FUNCTION_BLOCK SortingRouteConditions (* Sorting-only architecture following Distribution and tutorial modules 1-4 *)
  (* Standard: 61499-2 *)
  (* Version 2.0, 2026-11-09, sorting2n, sorting2n *)
  PACKAGE Main;
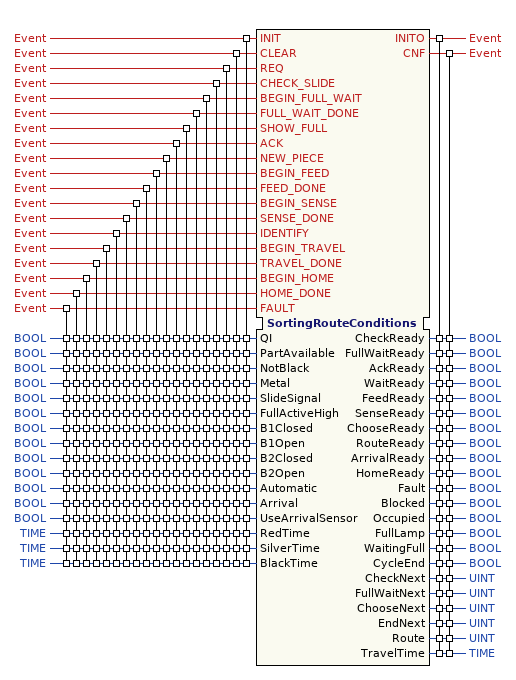
  EVENT_INPUT
    INIT WITH QI, PartAvailable, NotBlack, Metal, SlideSignal, FullActiveHigh, B1Closed, B1Open, B2Closed, B2Open, Automatic, Arrival, UseArrivalSensor, RedTime, SilverTime, BlackTime;
    CLEAR WITH QI, PartAvailable, NotBlack, Metal, SlideSignal, FullActiveHigh, B1Closed, B1Open, B2Closed, B2Open, Automatic, Arrival, UseArrivalSensor, RedTime, SilverTime, BlackTime;
    REQ WITH QI, PartAvailable, NotBlack, Metal, SlideSignal, FullActiveHigh, B1Closed, B1Open, B2Closed, B2Open, Automatic, Arrival, UseArrivalSensor, RedTime, SilverTime, BlackTime;
    CHECK_SLIDE WITH QI, PartAvailable, NotBlack, Metal, SlideSignal, FullActiveHigh, B1Closed, B1Open, B2Closed, B2Open, Automatic, Arrival, UseArrivalSensor, RedTime, SilverTime, BlackTime;
    BEGIN_FULL_WAIT WITH QI, PartAvailable, NotBlack, Metal, SlideSignal, FullActiveHigh, B1Closed, B1Open, B2Closed, B2Open, Automatic, Arrival, UseArrivalSensor, RedTime, SilverTime, BlackTime;
    FULL_WAIT_DONE WITH QI, PartAvailable, NotBlack, Metal, SlideSignal, FullActiveHigh, B1Closed, B1Open, B2Closed, B2Open, Automatic, Arrival, UseArrivalSensor, RedTime, SilverTime, BlackTime;
    SHOW_FULL WITH QI, PartAvailable, NotBlack, Metal, SlideSignal, FullActiveHigh, B1Closed, B1Open, B2Closed, B2Open, Automatic, Arrival, UseArrivalSensor, RedTime, SilverTime, BlackTime;
    ACK WITH QI, PartAvailable, NotBlack, Metal, SlideSignal, FullActiveHigh, B1Closed, B1Open, B2Closed, B2Open, Automatic, Arrival, UseArrivalSensor, RedTime, SilverTime, BlackTime;
    NEW_PIECE WITH QI, PartAvailable, NotBlack, Metal, SlideSignal, FullActiveHigh, B1Closed, B1Open, B2Closed, B2Open, Automatic, Arrival, UseArrivalSensor, RedTime, SilverTime, BlackTime;
    BEGIN_FEED WITH QI, PartAvailable, NotBlack, Metal, SlideSignal, FullActiveHigh, B1Closed, B1Open, B2Closed, B2Open, Automatic, Arrival, UseArrivalSensor, RedTime, SilverTime, BlackTime;
    FEED_DONE WITH QI, PartAvailable, NotBlack, Metal, SlideSignal, FullActiveHigh, B1Closed, B1Open, B2Closed, B2Open, Automatic, Arrival, UseArrivalSensor, RedTime, SilverTime, BlackTime;
    BEGIN_SENSE WITH QI, PartAvailable, NotBlack, Metal, SlideSignal, FullActiveHigh, B1Closed, B1Open, B2Closed, B2Open, Automatic, Arrival, UseArrivalSensor, RedTime, SilverTime, BlackTime;
    SENSE_DONE WITH QI, PartAvailable, NotBlack, Metal, SlideSignal, FullActiveHigh, B1Closed, B1Open, B2Closed, B2Open, Automatic, Arrival, UseArrivalSensor, RedTime, SilverTime, BlackTime;
    IDENTIFY WITH QI, PartAvailable, NotBlack, Metal, SlideSignal, FullActiveHigh, B1Closed, B1Open, B2Closed, B2Open, Automatic, Arrival, UseArrivalSensor, RedTime, SilverTime, BlackTime;
    BEGIN_TRAVEL WITH QI, PartAvailable, NotBlack, Metal, SlideSignal, FullActiveHigh, B1Closed, B1Open, B2Closed, B2Open, Automatic, Arrival, UseArrivalSensor, RedTime, SilverTime, BlackTime;
    TRAVEL_DONE WITH QI, PartAvailable, NotBlack, Metal, SlideSignal, FullActiveHigh, B1Closed, B1Open, B2Closed, B2Open, Automatic, Arrival, UseArrivalSensor, RedTime, SilverTime, BlackTime;
    BEGIN_HOME WITH QI, PartAvailable, NotBlack, Metal, SlideSignal, FullActiveHigh, B1Closed, B1Open, B2Closed, B2Open, Automatic, Arrival, UseArrivalSensor, RedTime, SilverTime, BlackTime;
    HOME_DONE WITH QI, PartAvailable, NotBlack, Metal, SlideSignal, FullActiveHigh, B1Closed, B1Open, B2Closed, B2Open, Automatic, Arrival, UseArrivalSensor, RedTime, SilverTime, BlackTime;
    FAULT WITH QI, PartAvailable, NotBlack, Metal, SlideSignal, FullActiveHigh, B1Closed, B1Open, B2Closed, B2Open, Automatic, Arrival, UseArrivalSensor, RedTime, SilverTime, BlackTime;
  END_EVENT
  EVENT_OUTPUT
    INITO WITH CheckReady, FullWaitReady, AckReady, WaitReady, FeedReady, SenseReady, ChooseReady, RouteReady, ArrivalReady, HomeReady, Fault, Blocked, Occupied, FullLamp, WaitingFull, CycleEnd, CheckNext, FullWaitNext, ChooseNext, EndNext, Route, TravelTime;
    CNF WITH CheckReady, FullWaitReady, AckReady, WaitReady, FeedReady, SenseReady, ChooseReady, RouteReady, ArrivalReady, HomeReady, Fault, Blocked, Occupied, FullLamp, WaitingFull, CycleEnd, CheckNext, FullWaitNext, ChooseNext, EndNext, Route, TravelTime;
  END_EVENT
  VAR_INPUT
    QI : BOOL := FALSE;
    PartAvailable : BOOL := FALSE;
    NotBlack : BOOL := FALSE;
    Metal : BOOL := FALSE;
    SlideSignal : BOOL := FALSE;
    FullActiveHigh : BOOL := FALSE;
    B1Closed : BOOL := FALSE;
    B1Open : BOOL := FALSE;
    B2Closed : BOOL := FALSE;
    B2Open : BOOL := FALSE;
    Automatic : BOOL := FALSE;
    Arrival : BOOL := FALSE;
    UseArrivalSensor : BOOL := FALSE;
    RedTime : TIME := T#2500ms;
    SilverTime : TIME := T#3s;
    BlackTime : TIME := T#5s;
  END_VAR
  VAR_OUTPUT
    CheckReady : BOOL := FALSE;
    FullWaitReady : BOOL := FALSE;
    AckReady : BOOL := FALSE;
    WaitReady : BOOL := FALSE;
    FeedReady : BOOL := FALSE;
    SenseReady : BOOL := FALSE;
    ChooseReady : BOOL := FALSE;
    RouteReady : BOOL := FALSE;
    ArrivalReady : BOOL := FALSE;
    HomeReady : BOOL := FALSE;
    Fault : BOOL := FALSE;
    Blocked : BOOL := FALSE;
    Occupied : BOOL := FALSE;
    FullLamp : BOOL := FALSE;
    WaitingFull : BOOL := FALSE;
    CycleEnd : BOOL := FALSE;
    CheckNext : UINT := 0;
    FullWaitNext : UINT := 0;
    ChooseNext : UINT := 0;
    EndNext : UINT := 0;
    Route : UINT := 0;
    TravelTime : TIME := T#5s;
  END_VAR
  VAR
    FeedElapsed : BOOL;
    SenseElapsed : BOOL;
    FinishElapsed : BOOL;
    TravelElapsed : BOOL;
    HomeElapsed : BOOL;
    Acked : BOOL;
  END_VAR
  EC_STATES
    IDLE;
    ON_INIT : ON_INIT -> INITO;
    ON_CLEAR : ON_CLEAR -> CNF;
    ON_REQ : ON_REQ -> CNF;
    ON_CHECK_SLIDE : ON_CHECK_SLIDE -> CNF;
    ON_BEGIN_FULL_WAIT : ON_BEGIN_FULL_WAIT -> CNF;
    ON_FULL_WAIT_DONE : ON_FULL_WAIT_DONE -> CNF;
    ON_SHOW_FULL : ON_SHOW_FULL -> CNF;
    ON_ACK : ON_ACK -> CNF;
    ON_NEW_PIECE : ON_NEW_PIECE -> CNF;
    ON_BEGIN_FEED : ON_BEGIN_FEED -> CNF;
    ON_FEED_DONE : ON_FEED_DONE -> CNF;
    ON_BEGIN_SENSE : ON_BEGIN_SENSE -> CNF;
    ON_SENSE_DONE : ON_SENSE_DONE -> CNF;
    ON_IDENTIFY : ON_IDENTIFY -> CNF;
    ON_BEGIN_TRAVEL : ON_BEGIN_TRAVEL -> CNF;
    ON_TRAVEL_DONE : ON_TRAVEL_DONE -> CNF;
    ON_BEGIN_HOME : ON_BEGIN_HOME -> CNF;
    ON_HOME_DONE : ON_HOME_DONE -> CNF;
    ON_FAULT : ON_FAULT -> CNF;
  END_STATES
  EC_TRANSITIONS
    IDLE TO ON_INIT := INIT;
    ON_INIT TO IDLE := 1;
    IDLE TO ON_CLEAR := CLEAR;
    ON_CLEAR TO IDLE := 1;
    IDLE TO ON_REQ := REQ;
    ON_REQ TO IDLE := 1;
    IDLE TO ON_CHECK_SLIDE := CHECK_SLIDE;
    ON_CHECK_SLIDE TO IDLE := 1;
    IDLE TO ON_BEGIN_FULL_WAIT := BEGIN_FULL_WAIT;
    ON_BEGIN_FULL_WAIT TO IDLE := 1;
    IDLE TO ON_FULL_WAIT_DONE := FULL_WAIT_DONE;
    ON_FULL_WAIT_DONE TO IDLE := 1;
    IDLE TO ON_SHOW_FULL := SHOW_FULL;
    ON_SHOW_FULL TO IDLE := 1;
    IDLE TO ON_ACK := ACK;
    ON_ACK TO IDLE := 1;
    IDLE TO ON_NEW_PIECE := NEW_PIECE;
    ON_NEW_PIECE TO IDLE := 1;
    IDLE TO ON_BEGIN_FEED := BEGIN_FEED;
    ON_BEGIN_FEED TO IDLE := 1;
    IDLE TO ON_FEED_DONE := FEED_DONE;
    ON_FEED_DONE TO IDLE := 1;
    IDLE TO ON_BEGIN_SENSE := BEGIN_SENSE;
    ON_BEGIN_SENSE TO IDLE := 1;
    IDLE TO ON_SENSE_DONE := SENSE_DONE;
    ON_SENSE_DONE TO IDLE := 1;
    IDLE TO ON_IDENTIFY := IDENTIFY;
    ON_IDENTIFY TO IDLE := 1;
    IDLE TO ON_BEGIN_TRAVEL := BEGIN_TRAVEL;
    ON_BEGIN_TRAVEL TO IDLE := 1;
    IDLE TO ON_TRAVEL_DONE := TRAVEL_DONE;
    ON_TRAVEL_DONE TO IDLE := 1;
    IDLE TO ON_BEGIN_HOME := BEGIN_HOME;
    ON_BEGIN_HOME TO IDLE := 1;
    IDLE TO ON_HOME_DONE := HOME_DONE;
    ON_HOME_DONE TO IDLE := 1;
    IDLE TO ON_FAULT := FAULT;
    ON_FAULT TO IDLE := 1;
  END_TRANSITIONS
  ALGORITHM ON_INIT IN ST:
FeedElapsed := FALSE; SenseElapsed := FALSE; FinishElapsed := FALSE; TravelElapsed := FALSE; HomeElapsed := FALSE; Acked := FALSE; Route := 0; Fault := FALSE; Occupied := FALSE; FullLamp := FALSE; WaitingFull := FALSE; CycleEnd := FALSE;
IF FullActiveHigh THEN Blocked := SlideSignal; ELSE Blocked := NOT SlideSignal; END_IF;
IF (B1Closed AND B1Open) OR (B2Closed AND B2Open) THEN Fault := TRUE; END_IF;
CheckReady := QI AND NOT Fault; IF Blocked THEN CheckNext := 3; ELSE CheckNext := 5; END_IF;
FullWaitReady := FinishElapsed AND NOT Fault; IF Blocked THEN FullWaitNext := 4; ELSE FullWaitNext := 2; END_IF;
AckReady := Acked AND NOT Fault;
WaitReady := QI AND PartAvailable AND NOT Fault;
FeedReady := FeedElapsed AND NOT PartAvailable AND NOT Fault;
SenseReady := SenseElapsed AND NOT Fault;
ChooseReady := (Route > 0) AND NOT Fault;
IF Route = 1 THEN ChooseNext := 9; ELSIF Route = 2 THEN ChooseNext := 11; ELSE ChooseNext := 13; END_IF;
RouteReady := ChooseReady AND ((Route = 1 AND B1Open AND B2Closed) OR (Route = 2 AND B1Closed AND B2Open) OR (Route = 3 AND B1Closed AND B2Closed));
ArrivalReady := ((UseArrivalSensor AND Arrival) OR (NOT UseArrivalSensor AND TravelElapsed)) AND NOT Fault;
HomeReady := HomeElapsed AND B1Closed AND B2Closed AND NOT Fault;
IF Automatic THEN EndNext := 2; ELSE EndNext := 15; END_IF;
TravelTime := BlackTime; IF Route = 1 THEN TravelTime := RedTime; ELSIF Route = 2 THEN TravelTime := SilverTime; END_IF;
  END_ALGORITHM
  ALGORITHM ON_CLEAR IN ST:
FeedElapsed := FALSE; SenseElapsed := FALSE; FinishElapsed := FALSE; TravelElapsed := FALSE; HomeElapsed := FALSE; Acked := FALSE; Route := 0; Fault := FALSE; Occupied := FALSE; FullLamp := FALSE; WaitingFull := FALSE; CycleEnd := FALSE;
IF FullActiveHigh THEN Blocked := SlideSignal; ELSE Blocked := NOT SlideSignal; END_IF;
IF (B1Closed AND B1Open) OR (B2Closed AND B2Open) THEN Fault := TRUE; END_IF;
CheckReady := QI AND NOT Fault; IF Blocked THEN CheckNext := 3; ELSE CheckNext := 5; END_IF;
FullWaitReady := FinishElapsed AND NOT Fault; IF Blocked THEN FullWaitNext := 4; ELSE FullWaitNext := 2; END_IF;
AckReady := Acked AND NOT Fault;
WaitReady := QI AND PartAvailable AND NOT Fault;
FeedReady := FeedElapsed AND NOT PartAvailable AND NOT Fault;
SenseReady := SenseElapsed AND NOT Fault;
ChooseReady := (Route > 0) AND NOT Fault;
IF Route = 1 THEN ChooseNext := 9; ELSIF Route = 2 THEN ChooseNext := 11; ELSE ChooseNext := 13; END_IF;
RouteReady := ChooseReady AND ((Route = 1 AND B1Open AND B2Closed) OR (Route = 2 AND B1Closed AND B2Open) OR (Route = 3 AND B1Closed AND B2Closed));
ArrivalReady := ((UseArrivalSensor AND Arrival) OR (NOT UseArrivalSensor AND TravelElapsed)) AND NOT Fault;
HomeReady := HomeElapsed AND B1Closed AND B2Closed AND NOT Fault;
IF Automatic THEN EndNext := 2; ELSE EndNext := 15; END_IF;
TravelTime := BlackTime; IF Route = 1 THEN TravelTime := RedTime; ELSIF Route = 2 THEN TravelTime := SilverTime; END_IF;
  END_ALGORITHM
  ALGORITHM ON_REQ IN ST:
IF FullActiveHigh THEN Blocked := SlideSignal; ELSE Blocked := NOT SlideSignal; END_IF;
IF (B1Closed AND B1Open) OR (B2Closed AND B2Open) THEN Fault := TRUE; END_IF;
CheckReady := QI AND NOT Fault; IF Blocked THEN CheckNext := 3; ELSE CheckNext := 5; END_IF;
FullWaitReady := FinishElapsed AND NOT Fault; IF Blocked THEN FullWaitNext := 4; ELSE FullWaitNext := 2; END_IF;
AckReady := Acked AND NOT Fault;
WaitReady := QI AND PartAvailable AND NOT Fault;
FeedReady := FeedElapsed AND NOT PartAvailable AND NOT Fault;
SenseReady := SenseElapsed AND NOT Fault;
ChooseReady := (Route > 0) AND NOT Fault;
IF Route = 1 THEN ChooseNext := 9; ELSIF Route = 2 THEN ChooseNext := 11; ELSE ChooseNext := 13; END_IF;
RouteReady := ChooseReady AND ((Route = 1 AND B1Open AND B2Closed) OR (Route = 2 AND B1Closed AND B2Open) OR (Route = 3 AND B1Closed AND B2Closed));
ArrivalReady := ((UseArrivalSensor AND Arrival) OR (NOT UseArrivalSensor AND TravelElapsed)) AND NOT Fault;
HomeReady := HomeElapsed AND B1Closed AND B2Closed AND NOT Fault;
IF Automatic THEN EndNext := 2; ELSE EndNext := 15; END_IF;
TravelTime := BlackTime; IF Route = 1 THEN TravelTime := RedTime; ELSIF Route = 2 THEN TravelTime := SilverTime; END_IF;
  END_ALGORITHM
  ALGORITHM ON_CHECK_SLIDE IN ST:
FullLamp := FALSE; WaitingFull := FALSE; CycleEnd := FALSE; IF FullActiveHigh THEN Blocked := SlideSignal; ELSE Blocked := NOT SlideSignal; END_IF; IF NOT Blocked THEN Occupied := FALSE; END_IF;
IF FullActiveHigh THEN Blocked := SlideSignal; ELSE Blocked := NOT SlideSignal; END_IF;
IF (B1Closed AND B1Open) OR (B2Closed AND B2Open) THEN Fault := TRUE; END_IF;
CheckReady := QI AND NOT Fault; IF Blocked THEN CheckNext := 3; ELSE CheckNext := 5; END_IF;
FullWaitReady := FinishElapsed AND NOT Fault; IF Blocked THEN FullWaitNext := 4; ELSE FullWaitNext := 2; END_IF;
AckReady := Acked AND NOT Fault;
WaitReady := QI AND PartAvailable AND NOT Fault;
FeedReady := FeedElapsed AND NOT PartAvailable AND NOT Fault;
SenseReady := SenseElapsed AND NOT Fault;
ChooseReady := (Route > 0) AND NOT Fault;
IF Route = 1 THEN ChooseNext := 9; ELSIF Route = 2 THEN ChooseNext := 11; ELSE ChooseNext := 13; END_IF;
RouteReady := ChooseReady AND ((Route = 1 AND B1Open AND B2Closed) OR (Route = 2 AND B1Closed AND B2Open) OR (Route = 3 AND B1Closed AND B2Closed));
ArrivalReady := ((UseArrivalSensor AND Arrival) OR (NOT UseArrivalSensor AND TravelElapsed)) AND NOT Fault;
HomeReady := HomeElapsed AND B1Closed AND B2Closed AND NOT Fault;
IF Automatic THEN EndNext := 2; ELSE EndNext := 15; END_IF;
TravelTime := BlackTime; IF Route = 1 THEN TravelTime := RedTime; ELSIF Route = 2 THEN TravelTime := SilverTime; END_IF;
  END_ALGORITHM
  ALGORITHM ON_BEGIN_FULL_WAIT IN ST:
FinishElapsed := FALSE;
IF FullActiveHigh THEN Blocked := SlideSignal; ELSE Blocked := NOT SlideSignal; END_IF;
IF (B1Closed AND B1Open) OR (B2Closed AND B2Open) THEN Fault := TRUE; END_IF;
CheckReady := QI AND NOT Fault; IF Blocked THEN CheckNext := 3; ELSE CheckNext := 5; END_IF;
FullWaitReady := FinishElapsed AND NOT Fault; IF Blocked THEN FullWaitNext := 4; ELSE FullWaitNext := 2; END_IF;
AckReady := Acked AND NOT Fault;
WaitReady := QI AND PartAvailable AND NOT Fault;
FeedReady := FeedElapsed AND NOT PartAvailable AND NOT Fault;
SenseReady := SenseElapsed AND NOT Fault;
ChooseReady := (Route > 0) AND NOT Fault;
IF Route = 1 THEN ChooseNext := 9; ELSIF Route = 2 THEN ChooseNext := 11; ELSE ChooseNext := 13; END_IF;
RouteReady := ChooseReady AND ((Route = 1 AND B1Open AND B2Closed) OR (Route = 2 AND B1Closed AND B2Open) OR (Route = 3 AND B1Closed AND B2Closed));
ArrivalReady := ((UseArrivalSensor AND Arrival) OR (NOT UseArrivalSensor AND TravelElapsed)) AND NOT Fault;
HomeReady := HomeElapsed AND B1Closed AND B2Closed AND NOT Fault;
IF Automatic THEN EndNext := 2; ELSE EndNext := 15; END_IF;
TravelTime := BlackTime; IF Route = 1 THEN TravelTime := RedTime; ELSIF Route = 2 THEN TravelTime := SilverTime; END_IF;
  END_ALGORITHM
  ALGORITHM ON_FULL_WAIT_DONE IN ST:
FinishElapsed := TRUE;
IF FullActiveHigh THEN Blocked := SlideSignal; ELSE Blocked := NOT SlideSignal; END_IF;
IF (B1Closed AND B1Open) OR (B2Closed AND B2Open) THEN Fault := TRUE; END_IF;
CheckReady := QI AND NOT Fault; IF Blocked THEN CheckNext := 3; ELSE CheckNext := 5; END_IF;
FullWaitReady := FinishElapsed AND NOT Fault; IF Blocked THEN FullWaitNext := 4; ELSE FullWaitNext := 2; END_IF;
AckReady := Acked AND NOT Fault;
WaitReady := QI AND PartAvailable AND NOT Fault;
FeedReady := FeedElapsed AND NOT PartAvailable AND NOT Fault;
SenseReady := SenseElapsed AND NOT Fault;
ChooseReady := (Route > 0) AND NOT Fault;
IF Route = 1 THEN ChooseNext := 9; ELSIF Route = 2 THEN ChooseNext := 11; ELSE ChooseNext := 13; END_IF;
RouteReady := ChooseReady AND ((Route = 1 AND B1Open AND B2Closed) OR (Route = 2 AND B1Closed AND B2Open) OR (Route = 3 AND B1Closed AND B2Closed));
ArrivalReady := ((UseArrivalSensor AND Arrival) OR (NOT UseArrivalSensor AND TravelElapsed)) AND NOT Fault;
HomeReady := HomeElapsed AND B1Closed AND B2Closed AND NOT Fault;
IF Automatic THEN EndNext := 2; ELSE EndNext := 15; END_IF;
TravelTime := BlackTime; IF Route = 1 THEN TravelTime := RedTime; ELSIF Route = 2 THEN TravelTime := SilverTime; END_IF;
  END_ALGORITHM
  ALGORITHM ON_SHOW_FULL IN ST:
Occupied := TRUE; FullLamp := TRUE; WaitingFull := TRUE; Acked := FALSE;
IF FullActiveHigh THEN Blocked := SlideSignal; ELSE Blocked := NOT SlideSignal; END_IF;
IF (B1Closed AND B1Open) OR (B2Closed AND B2Open) THEN Fault := TRUE; END_IF;
CheckReady := QI AND NOT Fault; IF Blocked THEN CheckNext := 3; ELSE CheckNext := 5; END_IF;
FullWaitReady := FinishElapsed AND NOT Fault; IF Blocked THEN FullWaitNext := 4; ELSE FullWaitNext := 2; END_IF;
AckReady := Acked AND NOT Fault;
WaitReady := QI AND PartAvailable AND NOT Fault;
FeedReady := FeedElapsed AND NOT PartAvailable AND NOT Fault;
SenseReady := SenseElapsed AND NOT Fault;
ChooseReady := (Route > 0) AND NOT Fault;
IF Route = 1 THEN ChooseNext := 9; ELSIF Route = 2 THEN ChooseNext := 11; ELSE ChooseNext := 13; END_IF;
RouteReady := ChooseReady AND ((Route = 1 AND B1Open AND B2Closed) OR (Route = 2 AND B1Closed AND B2Open) OR (Route = 3 AND B1Closed AND B2Closed));
ArrivalReady := ((UseArrivalSensor AND Arrival) OR (NOT UseArrivalSensor AND TravelElapsed)) AND NOT Fault;
HomeReady := HomeElapsed AND B1Closed AND B2Closed AND NOT Fault;
IF Automatic THEN EndNext := 2; ELSE EndNext := 15; END_IF;
TravelTime := BlackTime; IF Route = 1 THEN TravelTime := RedTime; ELSIF Route = 2 THEN TravelTime := SilverTime; END_IF;
  END_ALGORITHM
  ALGORITHM ON_ACK IN ST:
Acked := TRUE;
IF FullActiveHigh THEN Blocked := SlideSignal; ELSE Blocked := NOT SlideSignal; END_IF;
IF (B1Closed AND B1Open) OR (B2Closed AND B2Open) THEN Fault := TRUE; END_IF;
CheckReady := QI AND NOT Fault; IF Blocked THEN CheckNext := 3; ELSE CheckNext := 5; END_IF;
FullWaitReady := FinishElapsed AND NOT Fault; IF Blocked THEN FullWaitNext := 4; ELSE FullWaitNext := 2; END_IF;
AckReady := Acked AND NOT Fault;
WaitReady := QI AND PartAvailable AND NOT Fault;
FeedReady := FeedElapsed AND NOT PartAvailable AND NOT Fault;
SenseReady := SenseElapsed AND NOT Fault;
ChooseReady := (Route > 0) AND NOT Fault;
IF Route = 1 THEN ChooseNext := 9; ELSIF Route = 2 THEN ChooseNext := 11; ELSE ChooseNext := 13; END_IF;
RouteReady := ChooseReady AND ((Route = 1 AND B1Open AND B2Closed) OR (Route = 2 AND B1Closed AND B2Open) OR (Route = 3 AND B1Closed AND B2Closed));
ArrivalReady := ((UseArrivalSensor AND Arrival) OR (NOT UseArrivalSensor AND TravelElapsed)) AND NOT Fault;
HomeReady := HomeElapsed AND B1Closed AND B2Closed AND NOT Fault;
IF Automatic THEN EndNext := 2; ELSE EndNext := 15; END_IF;
TravelTime := BlackTime; IF Route = 1 THEN TravelTime := RedTime; ELSIF Route = 2 THEN TravelTime := SilverTime; END_IF;
  END_ALGORITHM
  ALGORITHM ON_NEW_PIECE IN ST:
Route := 0; FeedElapsed := FALSE; SenseElapsed := FALSE; TravelElapsed := FALSE; HomeElapsed := FALSE; Occupied := FALSE; CycleEnd := FALSE;
IF FullActiveHigh THEN Blocked := SlideSignal; ELSE Blocked := NOT SlideSignal; END_IF;
IF (B1Closed AND B1Open) OR (B2Closed AND B2Open) THEN Fault := TRUE; END_IF;
CheckReady := QI AND NOT Fault; IF Blocked THEN CheckNext := 3; ELSE CheckNext := 5; END_IF;
FullWaitReady := FinishElapsed AND NOT Fault; IF Blocked THEN FullWaitNext := 4; ELSE FullWaitNext := 2; END_IF;
AckReady := Acked AND NOT Fault;
WaitReady := QI AND PartAvailable AND NOT Fault;
FeedReady := FeedElapsed AND NOT PartAvailable AND NOT Fault;
SenseReady := SenseElapsed AND NOT Fault;
ChooseReady := (Route > 0) AND NOT Fault;
IF Route = 1 THEN ChooseNext := 9; ELSIF Route = 2 THEN ChooseNext := 11; ELSE ChooseNext := 13; END_IF;
RouteReady := ChooseReady AND ((Route = 1 AND B1Open AND B2Closed) OR (Route = 2 AND B1Closed AND B2Open) OR (Route = 3 AND B1Closed AND B2Closed));
ArrivalReady := ((UseArrivalSensor AND Arrival) OR (NOT UseArrivalSensor AND TravelElapsed)) AND NOT Fault;
HomeReady := HomeElapsed AND B1Closed AND B2Closed AND NOT Fault;
IF Automatic THEN EndNext := 2; ELSE EndNext := 15; END_IF;
TravelTime := BlackTime; IF Route = 1 THEN TravelTime := RedTime; ELSIF Route = 2 THEN TravelTime := SilverTime; END_IF;
  END_ALGORITHM
  ALGORITHM ON_BEGIN_FEED IN ST:
FeedElapsed := FALSE; Occupied := TRUE;
IF FullActiveHigh THEN Blocked := SlideSignal; ELSE Blocked := NOT SlideSignal; END_IF;
IF (B1Closed AND B1Open) OR (B2Closed AND B2Open) THEN Fault := TRUE; END_IF;
CheckReady := QI AND NOT Fault; IF Blocked THEN CheckNext := 3; ELSE CheckNext := 5; END_IF;
FullWaitReady := FinishElapsed AND NOT Fault; IF Blocked THEN FullWaitNext := 4; ELSE FullWaitNext := 2; END_IF;
AckReady := Acked AND NOT Fault;
WaitReady := QI AND PartAvailable AND NOT Fault;
FeedReady := FeedElapsed AND NOT PartAvailable AND NOT Fault;
SenseReady := SenseElapsed AND NOT Fault;
ChooseReady := (Route > 0) AND NOT Fault;
IF Route = 1 THEN ChooseNext := 9; ELSIF Route = 2 THEN ChooseNext := 11; ELSE ChooseNext := 13; END_IF;
RouteReady := ChooseReady AND ((Route = 1 AND B1Open AND B2Closed) OR (Route = 2 AND B1Closed AND B2Open) OR (Route = 3 AND B1Closed AND B2Closed));
ArrivalReady := ((UseArrivalSensor AND Arrival) OR (NOT UseArrivalSensor AND TravelElapsed)) AND NOT Fault;
HomeReady := HomeElapsed AND B1Closed AND B2Closed AND NOT Fault;
IF Automatic THEN EndNext := 2; ELSE EndNext := 15; END_IF;
TravelTime := BlackTime; IF Route = 1 THEN TravelTime := RedTime; ELSIF Route = 2 THEN TravelTime := SilverTime; END_IF;
  END_ALGORITHM
  ALGORITHM ON_FEED_DONE IN ST:
FeedElapsed := TRUE;
IF FullActiveHigh THEN Blocked := SlideSignal; ELSE Blocked := NOT SlideSignal; END_IF;
IF (B1Closed AND B1Open) OR (B2Closed AND B2Open) THEN Fault := TRUE; END_IF;
CheckReady := QI AND NOT Fault; IF Blocked THEN CheckNext := 3; ELSE CheckNext := 5; END_IF;
FullWaitReady := FinishElapsed AND NOT Fault; IF Blocked THEN FullWaitNext := 4; ELSE FullWaitNext := 2; END_IF;
AckReady := Acked AND NOT Fault;
WaitReady := QI AND PartAvailable AND NOT Fault;
FeedReady := FeedElapsed AND NOT PartAvailable AND NOT Fault;
SenseReady := SenseElapsed AND NOT Fault;
ChooseReady := (Route > 0) AND NOT Fault;
IF Route = 1 THEN ChooseNext := 9; ELSIF Route = 2 THEN ChooseNext := 11; ELSE ChooseNext := 13; END_IF;
RouteReady := ChooseReady AND ((Route = 1 AND B1Open AND B2Closed) OR (Route = 2 AND B1Closed AND B2Open) OR (Route = 3 AND B1Closed AND B2Closed));
ArrivalReady := ((UseArrivalSensor AND Arrival) OR (NOT UseArrivalSensor AND TravelElapsed)) AND NOT Fault;
HomeReady := HomeElapsed AND B1Closed AND B2Closed AND NOT Fault;
IF Automatic THEN EndNext := 2; ELSE EndNext := 15; END_IF;
TravelTime := BlackTime; IF Route = 1 THEN TravelTime := RedTime; ELSIF Route = 2 THEN TravelTime := SilverTime; END_IF;
  END_ALGORITHM
  ALGORITHM ON_BEGIN_SENSE IN ST:
SenseElapsed := FALSE;
IF FullActiveHigh THEN Blocked := SlideSignal; ELSE Blocked := NOT SlideSignal; END_IF;
IF (B1Closed AND B1Open) OR (B2Closed AND B2Open) THEN Fault := TRUE; END_IF;
CheckReady := QI AND NOT Fault; IF Blocked THEN CheckNext := 3; ELSE CheckNext := 5; END_IF;
FullWaitReady := FinishElapsed AND NOT Fault; IF Blocked THEN FullWaitNext := 4; ELSE FullWaitNext := 2; END_IF;
AckReady := Acked AND NOT Fault;
WaitReady := QI AND PartAvailable AND NOT Fault;
FeedReady := FeedElapsed AND NOT PartAvailable AND NOT Fault;
SenseReady := SenseElapsed AND NOT Fault;
ChooseReady := (Route > 0) AND NOT Fault;
IF Route = 1 THEN ChooseNext := 9; ELSIF Route = 2 THEN ChooseNext := 11; ELSE ChooseNext := 13; END_IF;
RouteReady := ChooseReady AND ((Route = 1 AND B1Open AND B2Closed) OR (Route = 2 AND B1Closed AND B2Open) OR (Route = 3 AND B1Closed AND B2Closed));
ArrivalReady := ((UseArrivalSensor AND Arrival) OR (NOT UseArrivalSensor AND TravelElapsed)) AND NOT Fault;
HomeReady := HomeElapsed AND B1Closed AND B2Closed AND NOT Fault;
IF Automatic THEN EndNext := 2; ELSE EndNext := 15; END_IF;
TravelTime := BlackTime; IF Route = 1 THEN TravelTime := RedTime; ELSIF Route = 2 THEN TravelTime := SilverTime; END_IF;
  END_ALGORITHM
  ALGORITHM ON_SENSE_DONE IN ST:
SenseElapsed := TRUE;
IF FullActiveHigh THEN Blocked := SlideSignal; ELSE Blocked := NOT SlideSignal; END_IF;
IF (B1Closed AND B1Open) OR (B2Closed AND B2Open) THEN Fault := TRUE; END_IF;
CheckReady := QI AND NOT Fault; IF Blocked THEN CheckNext := 3; ELSE CheckNext := 5; END_IF;
FullWaitReady := FinishElapsed AND NOT Fault; IF Blocked THEN FullWaitNext := 4; ELSE FullWaitNext := 2; END_IF;
AckReady := Acked AND NOT Fault;
WaitReady := QI AND PartAvailable AND NOT Fault;
FeedReady := FeedElapsed AND NOT PartAvailable AND NOT Fault;
SenseReady := SenseElapsed AND NOT Fault;
ChooseReady := (Route > 0) AND NOT Fault;
IF Route = 1 THEN ChooseNext := 9; ELSIF Route = 2 THEN ChooseNext := 11; ELSE ChooseNext := 13; END_IF;
RouteReady := ChooseReady AND ((Route = 1 AND B1Open AND B2Closed) OR (Route = 2 AND B1Closed AND B2Open) OR (Route = 3 AND B1Closed AND B2Closed));
ArrivalReady := ((UseArrivalSensor AND Arrival) OR (NOT UseArrivalSensor AND TravelElapsed)) AND NOT Fault;
HomeReady := HomeElapsed AND B1Closed AND B2Closed AND NOT Fault;
IF Automatic THEN EndNext := 2; ELSE EndNext := 15; END_IF;
TravelTime := BlackTime; IF Route = 1 THEN TravelTime := RedTime; ELSIF Route = 2 THEN TravelTime := SilverTime; END_IF;
  END_ALGORITHM
  ALGORITHM ON_IDENTIFY IN ST:
IF Metal AND NotBlack THEN Route := 2; ELSIF NotBlack AND NOT Metal THEN Route := 1; ELSIF NOT NotBlack AND NOT Metal THEN Route := 3; ELSE Route := 0; Fault := TRUE; END_IF;
IF FullActiveHigh THEN Blocked := SlideSignal; ELSE Blocked := NOT SlideSignal; END_IF;
IF (B1Closed AND B1Open) OR (B2Closed AND B2Open) THEN Fault := TRUE; END_IF;
CheckReady := QI AND NOT Fault; IF Blocked THEN CheckNext := 3; ELSE CheckNext := 5; END_IF;
FullWaitReady := FinishElapsed AND NOT Fault; IF Blocked THEN FullWaitNext := 4; ELSE FullWaitNext := 2; END_IF;
AckReady := Acked AND NOT Fault;
WaitReady := QI AND PartAvailable AND NOT Fault;
FeedReady := FeedElapsed AND NOT PartAvailable AND NOT Fault;
SenseReady := SenseElapsed AND NOT Fault;
ChooseReady := (Route > 0) AND NOT Fault;
IF Route = 1 THEN ChooseNext := 9; ELSIF Route = 2 THEN ChooseNext := 11; ELSE ChooseNext := 13; END_IF;
RouteReady := ChooseReady AND ((Route = 1 AND B1Open AND B2Closed) OR (Route = 2 AND B1Closed AND B2Open) OR (Route = 3 AND B1Closed AND B2Closed));
ArrivalReady := ((UseArrivalSensor AND Arrival) OR (NOT UseArrivalSensor AND TravelElapsed)) AND NOT Fault;
HomeReady := HomeElapsed AND B1Closed AND B2Closed AND NOT Fault;
IF Automatic THEN EndNext := 2; ELSE EndNext := 15; END_IF;
TravelTime := BlackTime; IF Route = 1 THEN TravelTime := RedTime; ELSIF Route = 2 THEN TravelTime := SilverTime; END_IF;
  END_ALGORITHM
  ALGORITHM ON_BEGIN_TRAVEL IN ST:
TravelElapsed := FALSE;
IF FullActiveHigh THEN Blocked := SlideSignal; ELSE Blocked := NOT SlideSignal; END_IF;
IF (B1Closed AND B1Open) OR (B2Closed AND B2Open) THEN Fault := TRUE; END_IF;
CheckReady := QI AND NOT Fault; IF Blocked THEN CheckNext := 3; ELSE CheckNext := 5; END_IF;
FullWaitReady := FinishElapsed AND NOT Fault; IF Blocked THEN FullWaitNext := 4; ELSE FullWaitNext := 2; END_IF;
AckReady := Acked AND NOT Fault;
WaitReady := QI AND PartAvailable AND NOT Fault;
FeedReady := FeedElapsed AND NOT PartAvailable AND NOT Fault;
SenseReady := SenseElapsed AND NOT Fault;
ChooseReady := (Route > 0) AND NOT Fault;
IF Route = 1 THEN ChooseNext := 9; ELSIF Route = 2 THEN ChooseNext := 11; ELSE ChooseNext := 13; END_IF;
RouteReady := ChooseReady AND ((Route = 1 AND B1Open AND B2Closed) OR (Route = 2 AND B1Closed AND B2Open) OR (Route = 3 AND B1Closed AND B2Closed));
ArrivalReady := ((UseArrivalSensor AND Arrival) OR (NOT UseArrivalSensor AND TravelElapsed)) AND NOT Fault;
HomeReady := HomeElapsed AND B1Closed AND B2Closed AND NOT Fault;
IF Automatic THEN EndNext := 2; ELSE EndNext := 15; END_IF;
TravelTime := BlackTime; IF Route = 1 THEN TravelTime := RedTime; ELSIF Route = 2 THEN TravelTime := SilverTime; END_IF;
  END_ALGORITHM
  ALGORITHM ON_TRAVEL_DONE IN ST:
TravelElapsed := TRUE;
IF FullActiveHigh THEN Blocked := SlideSignal; ELSE Blocked := NOT SlideSignal; END_IF;
IF (B1Closed AND B1Open) OR (B2Closed AND B2Open) THEN Fault := TRUE; END_IF;
CheckReady := QI AND NOT Fault; IF Blocked THEN CheckNext := 3; ELSE CheckNext := 5; END_IF;
FullWaitReady := FinishElapsed AND NOT Fault; IF Blocked THEN FullWaitNext := 4; ELSE FullWaitNext := 2; END_IF;
AckReady := Acked AND NOT Fault;
WaitReady := QI AND PartAvailable AND NOT Fault;
FeedReady := FeedElapsed AND NOT PartAvailable AND NOT Fault;
SenseReady := SenseElapsed AND NOT Fault;
ChooseReady := (Route > 0) AND NOT Fault;
IF Route = 1 THEN ChooseNext := 9; ELSIF Route = 2 THEN ChooseNext := 11; ELSE ChooseNext := 13; END_IF;
RouteReady := ChooseReady AND ((Route = 1 AND B1Open AND B2Closed) OR (Route = 2 AND B1Closed AND B2Open) OR (Route = 3 AND B1Closed AND B2Closed));
ArrivalReady := ((UseArrivalSensor AND Arrival) OR (NOT UseArrivalSensor AND TravelElapsed)) AND NOT Fault;
HomeReady := HomeElapsed AND B1Closed AND B2Closed AND NOT Fault;
IF Automatic THEN EndNext := 2; ELSE EndNext := 15; END_IF;
TravelTime := BlackTime; IF Route = 1 THEN TravelTime := RedTime; ELSIF Route = 2 THEN TravelTime := SilverTime; END_IF;
  END_ALGORITHM
  ALGORITHM ON_BEGIN_HOME IN ST:
HomeElapsed := FALSE; CycleEnd := TRUE;
IF FullActiveHigh THEN Blocked := SlideSignal; ELSE Blocked := NOT SlideSignal; END_IF;
IF (B1Closed AND B1Open) OR (B2Closed AND B2Open) THEN Fault := TRUE; END_IF;
CheckReady := QI AND NOT Fault; IF Blocked THEN CheckNext := 3; ELSE CheckNext := 5; END_IF;
FullWaitReady := FinishElapsed AND NOT Fault; IF Blocked THEN FullWaitNext := 4; ELSE FullWaitNext := 2; END_IF;
AckReady := Acked AND NOT Fault;
WaitReady := QI AND PartAvailable AND NOT Fault;
FeedReady := FeedElapsed AND NOT PartAvailable AND NOT Fault;
SenseReady := SenseElapsed AND NOT Fault;
ChooseReady := (Route > 0) AND NOT Fault;
IF Route = 1 THEN ChooseNext := 9; ELSIF Route = 2 THEN ChooseNext := 11; ELSE ChooseNext := 13; END_IF;
RouteReady := ChooseReady AND ((Route = 1 AND B1Open AND B2Closed) OR (Route = 2 AND B1Closed AND B2Open) OR (Route = 3 AND B1Closed AND B2Closed));
ArrivalReady := ((UseArrivalSensor AND Arrival) OR (NOT UseArrivalSensor AND TravelElapsed)) AND NOT Fault;
HomeReady := HomeElapsed AND B1Closed AND B2Closed AND NOT Fault;
IF Automatic THEN EndNext := 2; ELSE EndNext := 15; END_IF;
TravelTime := BlackTime; IF Route = 1 THEN TravelTime := RedTime; ELSIF Route = 2 THEN TravelTime := SilverTime; END_IF;
  END_ALGORITHM
  ALGORITHM ON_HOME_DONE IN ST:
HomeElapsed := TRUE;
IF FullActiveHigh THEN Blocked := SlideSignal; ELSE Blocked := NOT SlideSignal; END_IF;
IF (B1Closed AND B1Open) OR (B2Closed AND B2Open) THEN Fault := TRUE; END_IF;
CheckReady := QI AND NOT Fault; IF Blocked THEN CheckNext := 3; ELSE CheckNext := 5; END_IF;
FullWaitReady := FinishElapsed AND NOT Fault; IF Blocked THEN FullWaitNext := 4; ELSE FullWaitNext := 2; END_IF;
AckReady := Acked AND NOT Fault;
WaitReady := QI AND PartAvailable AND NOT Fault;
FeedReady := FeedElapsed AND NOT PartAvailable AND NOT Fault;
SenseReady := SenseElapsed AND NOT Fault;
ChooseReady := (Route > 0) AND NOT Fault;
IF Route = 1 THEN ChooseNext := 9; ELSIF Route = 2 THEN ChooseNext := 11; ELSE ChooseNext := 13; END_IF;
RouteReady := ChooseReady AND ((Route = 1 AND B1Open AND B2Closed) OR (Route = 2 AND B1Closed AND B2Open) OR (Route = 3 AND B1Closed AND B2Closed));
ArrivalReady := ((UseArrivalSensor AND Arrival) OR (NOT UseArrivalSensor AND TravelElapsed)) AND NOT Fault;
HomeReady := HomeElapsed AND B1Closed AND B2Closed AND NOT Fault;
IF Automatic THEN EndNext := 2; ELSE EndNext := 15; END_IF;
TravelTime := BlackTime; IF Route = 1 THEN TravelTime := RedTime; ELSIF Route = 2 THEN TravelTime := SilverTime; END_IF;
  END_ALGORITHM
  ALGORITHM ON_FAULT IN ST:
Fault := TRUE;
IF FullActiveHigh THEN Blocked := SlideSignal; ELSE Blocked := NOT SlideSignal; END_IF;
IF (B1Closed AND B1Open) OR (B2Closed AND B2Open) THEN Fault := TRUE; END_IF;
CheckReady := QI AND NOT Fault; IF Blocked THEN CheckNext := 3; ELSE CheckNext := 5; END_IF;
FullWaitReady := FinishElapsed AND NOT Fault; IF Blocked THEN FullWaitNext := 4; ELSE FullWaitNext := 2; END_IF;
AckReady := Acked AND NOT Fault;
WaitReady := QI AND PartAvailable AND NOT Fault;
FeedReady := FeedElapsed AND NOT PartAvailable AND NOT Fault;
SenseReady := SenseElapsed AND NOT Fault;
ChooseReady := (Route > 0) AND NOT Fault;
IF Route = 1 THEN ChooseNext := 9; ELSIF Route = 2 THEN ChooseNext := 11; ELSE ChooseNext := 13; END_IF;
RouteReady := ChooseReady AND ((Route = 1 AND B1Open AND B2Closed) OR (Route = 2 AND B1Closed AND B2Open) OR (Route = 3 AND B1Closed AND B2Closed));
ArrivalReady := ((UseArrivalSensor AND Arrival) OR (NOT UseArrivalSensor AND TravelElapsed)) AND NOT Fault;
HomeReady := HomeElapsed AND B1Closed AND B2Closed AND NOT Fault;
IF Automatic THEN EndNext := 2; ELSE EndNext := 15; END_IF;
TravelTime := BlackTime; IF Route = 1 THEN TravelTime := RedTime; ELSIF Route = 2 THEN TravelTime := SilverTime; END_IF;
  END_ALGORITHM
END_FUNCTION_BLOCK
